DATA_BLOCK "DB_Motor_Banderas"
{ S7_Optimized_Access := 'TRUE' }
VERSION : 0.1
NON_RETAIN
"FB_Motor_Banderas"

BEGIN

END_DATA_BLOCK

